(* Schneider Machine Expert - Basic project Taller2.txt, file version 2.9.0.0 *)
(* ProjectInformations: Name=Nuevo proyecto *)

HARDWARE
  Cpu 0: TM221CE40R
  EthernetConfiguration: NetworkName=M221, IpAllocationMode=FixedAddress, IpAddress=0.0.0.0, SubnetMask=0.0.0.0
  SerialLineConfiguration: Baud=Baud19200, Parity=ParityEven, DataBits=DataBits8, StopBits=StopBits1, PhysicalMedium=PhysicalMediumRs485, TransmissionMode=TransmissionModeModbusRtu, SlaveId=1, Addressing=SlaveAddressing
  MastTask: UsePeriodScanMode=false, PeriodScan=100
  FastTask: Period=255
  CpuBehavior: StartingMode=StartAsPreviousState, AutoSaveRamOnEeprom=true, WatchdogPeriod=250

SYMBOLS  (address, symbol, comment, settings)
  %TM2        [Preset=3, Base=OneSecond]
  %C1         [Preset=3]

POU Nuevo POU
  (* SectionNumber=1 *)

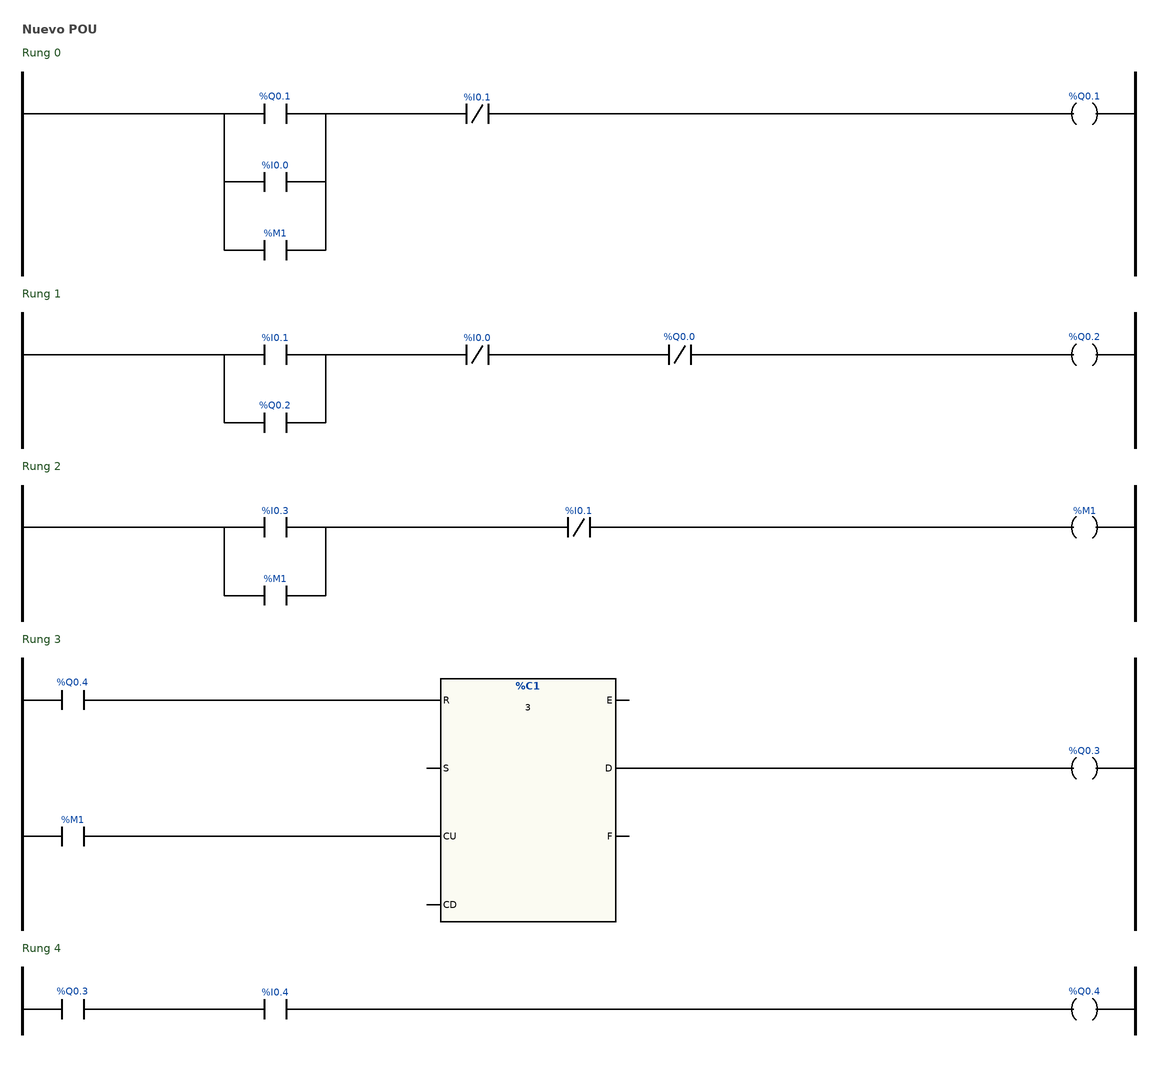

// Rung 0
  LD 1
  AND( %Q0.1
  OR %I0.0
  OR %M1
  )
  ANDN %I0.1
  ST %Q0.1
  // as ST:
  //   %Q0.1 := (%Q0.1 OR %I0.0 OR %M1) AND NOT %I0.1;

// Rung 1
  LD 1
  AND( %I0.1
  OR %Q0.2
  )
  ANDN %I0.0
  ANDN %Q0.0
  ST %Q0.2
  // as ST:
  //   %Q0.2 := (%I0.1 OR %Q0.2) AND NOT %I0.0 AND NOT %Q0.0;

// Rung 2
  LD 1
  AND( %I0.3
  OR %M1
  )
  ANDN %I0.1
  ST %M1
  // as ST:
  //   %M1 := (%I0.3 OR %M1) AND NOT %I0.1;

// Rung 3
  BLK %C1
  LD %Q0.4
  R
  LD %M1
  CU
  OUT_BLK
  LD D
  ST %Q0.3
  END_BLK
  // as ST:
  //   %C1(R := %Q0.4, CU := %M1);
  //   %Q0.3 := %C1.D;

// Rung 4
  LD %Q0.3
  AND %I0.4
  ST %Q0.4
  // as ST:
  //   %Q0.4 := %Q0.3 AND %I0.4;

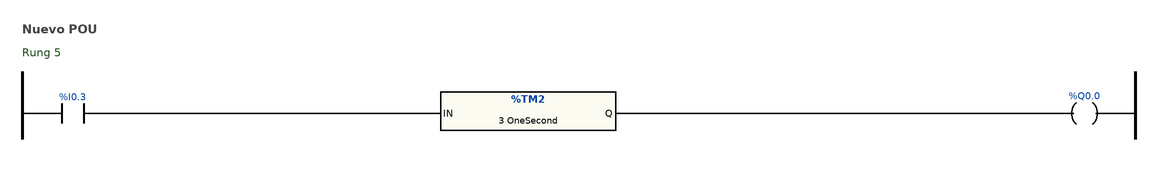

// Rung 5
  BLK %TM2
  LD %I0.3
  IN
  OUT_BLK
  LD Q
  ST %Q0.0
  END_BLK
  // as ST:
  //   %TM2(IN := %I0.3);
  //   %Q0.0 := %TM2.Q;
